(* IEC 61131-3 sources: kns-pump-station/tests/POUs/Station/FB_StationMode_Test, 10 files *)

(* ---- AutoToManualRequestsManual.method.decl.st ---- *)
// 04 §3.2: «Автомат» → «Ручной» — RequestMode(Manual) насосам в Auto и Local, OutOfService не трогается; событие
// 101002
METHOD PRIVATE AutoToManualRequestsManual
VAR
    fbDut    : FB_StationMode;                     // ФБ под тестом
    afbPump  : ARRAY[1..3] OF FB_FakeMotorVfd;     // подменные насосы
    fbSink   : FB_FakeEventSink;                   // подменный журнал
    stRetain : ST_StationRetain;                   // энергонезависимые данные станции
END_VAR

(* ---- EmptyRetainStartsManual.method.decl.st ---- *)
// 04 §3.2: пустой retain (умолчания типа) — станция в «Ручном», способ «Ступенчатое»; первый вызов даёт импульс
// входа в «Ручной» без запросов насосам и без событий
METHOD PRIVATE EmptyRetainStartsManual
VAR
    fbDut    : FB_StationMode;                     // ФБ под тестом
    afbPump  : ARRAY[1..3] OF FB_FakeMotorVfd;     // подменные насосы
    fbSink   : FB_FakeEventSink;                   // подменный журнал
    stRetain : ST_StationRetain;                   // энергонезависимые данные станции
END_VAR

(* ---- EnteredAutoPulsesOnFirstCallInAuto.method.decl.st ---- *)
// 04 §13.3: старт ПЛК с «Автоматом» в retain — импульс xEnteredAuto в первом вызове (подхват работающих насосов)
// без запросов режима и без события
METHOD PRIVATE EnteredAutoPulsesOnFirstCallInAuto
VAR
    fbDut    : FB_StationMode;                     // ФБ под тестом
    afbPump  : ARRAY[1..3] OF FB_FakeMotorVfd;     // подменные насосы
    fbSink   : FB_FakeEventSink;                   // подменный журнал
    stRetain : ST_StationRetain;                   // энергонезависимые данные станции
END_VAR

(* ---- GarbageRetainSanitized.method.decl.st ---- *)
// Правило L4 контракта: мусор в retain (режим 7, способ 0) заменяется «Ручным» и «Ступенчатым» сравнениями и
// записывается обратно
METHOD PRIVATE GarbageRetainSanitized
VAR
    fbDut    : FB_StationMode;                     // ФБ под тестом
    afbPump  : ARRAY[1..3] OF FB_FakeMotorVfd;     // подменные насосы
    fbSink   : FB_FakeEventSink;                   // подменный журнал
    stRetain : ST_StationRetain;                   // энергонезависимые данные станции
    pRaw    : POINTER TO INT;                      // запись числа вне перечисления
END_VAR

(* ---- LocalPumpGetsRememberedMode.method.decl.st ---- *)
// API 2.2, PMI-31: у насоса в Local запрос режима меняет запомненный дистанционный режим, сам режим остаётся Local
METHOD PRIVATE LocalPumpGetsRememberedMode
VAR
    fbDut    : FB_StationMode;                     // ФБ под тестом
    afbPump  : ARRAY[1..3] OF FB_FakeMotorVfd;     // подменные насосы
    fbSink   : FB_FakeEventSink;                   // подменный журнал
    stRetain : ST_StationRetain;                   // энергонезависимые данные станции
END_VAR

(* ---- ManualToAutoRequestsAutoExceptOos.method.decl.st ---- *)
// 04 §3.2, PMI-30: «Ручной» → «Автомат» — RequestMode(Auto) насосам в Manual и Local, OutOfService не трогается,
// насос в Auto — без запроса; событие 101001, импульс xEnteredAuto
METHOD PRIVATE ManualToAutoRequestsAutoExceptOos
VAR
    fbDut    : FB_StationMode;                     // ФБ под тестом
    afbPump  : ARRAY[1..3] OF FB_FakeMotorVfd;     // подменные насосы
    fbSink   : FB_FakeEventSink;                   // подменный журнал
    stRetain : ST_StationRetain;                   // энергонезависимые данные станции
END_VAR

(* ---- ManualWinsOverAutoSameCall.method.decl.st ---- *)
// 04 §19.2: xSetManual старше xSetAuto в одном вызове (безопасный вариант); оба импульса — обработанные команды
METHOD PRIVATE ManualWinsOverAutoSameCall
VAR
    fbDut    : FB_StationMode;                     // ФБ под тестом
    afbPump  : ARRAY[1..3] OF FB_FakeMotorVfd;     // подменные насосы
    fbSink   : FB_FakeEventSink;                   // подменный журнал
    stRetain : ST_StationRetain;                   // энергонезависимые данные станции
END_VAR

(* ---- MethodSwitchLoggedAndRetained.method.decl.st ---- *)
// 04 §3.2, PMI-07: смена способа — в retain и в журнал (101004, 101003); xSetStepped старше xSetLevelPid; способ
// не зависит от режима станции
METHOD PRIVATE MethodSwitchLoggedAndRetained
VAR
    fbDut    : FB_StationMode;                     // ФБ под тестом
    afbPump  : ARRAY[1..3] OF FB_FakeMotorVfd;     // подменные насосы
    fbSink   : FB_FakeEventSink;                   // подменный журнал
    stRetain : ST_StationRetain;                   // энергонезависимые данные станции
END_VAR

(* ---- NoEventSinkIsSafe.method.decl.st ---- *)
// Журнал не задан (itfEvents = 0) — переходы выполняются без обращения к журналу
METHOD PRIVATE NoEventSinkIsSafe
VAR
    fbDut    : FB_StationMode;                     // ФБ под тестом
    stRetain : ST_StationRetain;                   // энергонезависимые данные
END_VAR

(* ---- SameModeCommandAcceptedNoRequests.method.decl.st ---- *)
// Команда того же режима — Accepted без запросов насосам, без события и без импульса входа
METHOD PRIVATE SameModeCommandAcceptedNoRequests
VAR
    fbDut    : FB_StationMode;                     // ФБ под тестом
    afbPump  : ARRAY[1..3] OF FB_FakeMotorVfd;     // подменные насосы
    fbSink   : FB_FakeEventSink;                   // подменный журнал
    stRetain : ST_StationRetain;                   // энергонезависимые данные станции
END_VAR
